{region 'Documentation'}
(*!
<summary>Checks non-overlapping BYTE/WORD array token counts and independent array bounds.</summary>
<description>
Adjacent tokens count separately; overlapping candidates do not share elements.
Word patterns deliberately contain equal low bytes with different high bytes.
Oversized tokens and empty selected ranges are normal parameter errors, not
manufactured empty arrays or invalid references.
Independent scenarios occupy two calls: bound Reset, then evaluation.
ProcessAssertions checks each call before ProcessTests advances. Literal expected
results belong to SelectScenario, not to a copy of the production comparison.
The local capture is cleared before each call and checked in subject-call order.
FirstFailedScenario and FailedDuringEvaluation retain the first mismatch.
Continuation scenarios explicitly retain the prior subject state. The Test Case
owns all input storage; no invalid or dangling references are constructed.
</description>
*)
{endregion}
FUNCTION_BLOCK Test_AssertionArrayTokenCount EXTENDS TestCaseBase
VAR
    FEqual : AssertArrayTokenCntEqual_Byte;
    FEqualExpectedResult : E_Result;
    FWideEqual : AssertArrayTokenCntEqual_Word;
    FWideEqualExpectedResult : E_Result;
    FNone : AssertNoArrayToken_Byte;
    FNoneExpectedResult : E_Result;
    FWideRange : AssertArrayTokenCntInRange_Word;
    FWideRangeExpectedResult : E_Result;
    FData : ARRAY[-2..3] OF BYTE;
    FDataBefore : ARRAY[-2..3] OF BYTE;
    FWideData : ARRAY[-2..3] OF WORD;
    FWideDataBefore : ARRAY[-2..3] OF WORD;
    FToken : ARRAY[4..5] OF BYTE;
    FTokenBefore : ARRAY[4..5] OF BYTE;
    FWideToken : ARRAY[-5..-4] OF WORD;
    FWideTokenBefore : ARRAY[-5..-4] OF WORD;
    FStartIndex : DINT;
    FLength : USINT;
    FExpected : UINT;
    FMinimum : UINT;
    FMaximum : UINT;
    FSubjectEnable : BOOL;
    FContinueScenario : BOOL;
    FEqualExpectedFinding : BOOL;
    FEqualExpectedCount : UINT;
    FWideEqualExpectedFinding : BOOL;
    FWideEqualExpectedCount : UINT;
    FNoneExpectedFinding : BOOL;
    FNoneExpectedCount : UINT;
    FWideRangeExpectedFinding : BOOL;
    FWideRangeExpectedCount : UINT;
    FCapture : EventBuffer;
    FEvents : ARRAY[1..CaptureLength] OF ST_Event;
    FCaptureFifo : ST_FifoStatus;
    FCaptureStatus : ST_EventBufferStatus;
    FSetupValid : BOOL;
    FScenario : UINT;
    FChecked : BOOL;
    FEvaluateSubjects : BOOL;
    FObservationReady : BOOL;
    FFirstFailedScenario : UINT;
    FFailedDuringEvaluation : BOOL;
    FResultsMatch : BOOL;
    FResults : AssertTrue;
    FActivityMatch : BOOL;
    FActivity : AssertTrue;
    FInputsMatch : BOOL;
    FInputs : AssertTrue;
    FFindingsMatch : BOOL;
    FFindings : AssertTrue;
END_VAR
VAR CONSTANT
    CaptureLength : UINT := 8;
    ScenarioAdjacentTokens : UINT := 1;
    ScenarioNonOverlapping : UINT := 2;
    ScenarioTrailingPartial : UINT := 3;
    ScenarioLastCandidate : UINT := 4;
    ScenarioAbsent : UINT := 5;
    ScenarioCountMismatch : UINT := 6;
    ScenarioTokenTooLong : UINT := 7;
    ScenarioEmptyRange : UINT := 8;
    ScenarioRangePastEnd : UINT := 9;
    LastScenario : UINT := ScenarioRangePastEnd;
END_VAR

SUPER^();

{region 'Documentation'}
(*!
<summary>Aggregates only outer checks, not intentionally failing subjects.</summary>
*)
{endregion}
METHOD PROTECTED AggregateResults
VAR_INPUT
    Aggregator : I_ResultAggregator; //! Borrowed result sink owned by the outer Test Case; add this test's checking Assertions without resetting or retaining the sink.
END_VAR
Aggregator.AddProvider(Provider := FResults);
Aggregator.AddProvider(Provider := FActivity);
Aggregator.AddProvider(Provider := FInputs);
Aggregator.AddProvider(Provider := FFindings);
END_METHOD

{region 'Documentation'}
(*!
<summary>Calls each inherited production subject once with caller-owned input storage.</summary>
*)
{endregion}
METHOD PRIVATE CallSubjects
FEqual(Enable := FSubjectEnable,
    State := E_State.Running,
    StartIndex := FStartIndex,
    Length := FLength,
    Expected := FExpected,
    IN := FData,
    Token := FToken);
FWideEqual(Enable := FSubjectEnable,
    State := E_State.Running,
    StartIndex := FStartIndex,
    Length := FLength,
    Expected := FExpected,
    IN := FWideData,
    Token := FWideToken);
FNone(Enable := FSubjectEnable,
    State := E_State.Running,
    StartIndex := FStartIndex,
    Length := FLength,
    IN := FData,
    Token := FToken);
FWideRange(Enable := FSubjectEnable,
    State := E_State.Running,
    StartIndex := FStartIndex,
    Length := FLength,
    Minimum := FMinimum,
    Maximum := FMaximum,
    IN := FWideData,
    Token := FWideToken);
END_METHOD

{region 'Documentation'}
(*!
<summary>Checks one subject finding in call order; expected outcomes come from the scenario.</summary>
*)
{endregion}
METHOD PRIVATE CheckFinding : BOOL //! TRUE when the required finding checks pass; calls requiring no finding also succeed.
VAR_INPUT
    Subject : I_Assertion; //! Assertion interface supplying the expected finding identity.
    ExpectedResult : E_Result; //! Independently authored result expected in the captured finding.
    ExpectedFinding : BOOL; //! TRUE when this scenario requires a finding during active evaluation.
END_VAR
VAR_IN_OUT
    Index : UINT; //! One-based next finding index; advanced when this call checks a required finding.
END_VAR
CheckFinding := TRUE;
IF FEvaluateSubjects AND ExpectedFinding THEN
    CheckFinding := (FEvents[Index].SequenceId = UINT_TO_UDINT(Index))
        AND (FEvents[Index].Name = Subject.Name)
        AND (FEvents[Index].OwnerScope = E_OwnerScope.Assertion)
        AND (FEvents[Index].EventType = E_EventType.Result)
        AND (FEvents[Index].State = E_State.Running)
        AND (FEvents[Index].Result = ExpectedResult)
        AND (FEvents[Index].Message <> '');
    Index := Index + 1;
END_IF;
END_METHOD

{region 'Documentation'}
(*!
<summary>Checks exact finding count and identities; at most one finding per subject.</summary>
*)
{endregion}
METHOD PRIVATE CheckFindings
VAR
    Index : UINT;
    Matches : BOOL;
END_VAR
Index := 1;
FFindingsMatch := TRUE;
Matches := CheckFinding(Subject := FEqual,
    ExpectedResult := FEqualExpectedResult,
    ExpectedFinding := FEqualExpectedFinding,
    Index := Index);
FFindingsMatch := FFindingsMatch AND Matches;
Matches := CheckFinding(Subject := FWideEqual,
    ExpectedResult := FWideEqualExpectedResult,
    ExpectedFinding := FWideEqualExpectedFinding,
    Index := Index);
FFindingsMatch := FFindingsMatch AND Matches;
Matches := CheckFinding(Subject := FNone,
    ExpectedResult := FNoneExpectedResult,
    ExpectedFinding := FNoneExpectedFinding,
    Index := Index);
FFindingsMatch := FFindingsMatch AND Matches;
Matches := CheckFinding(Subject := FWideRange,
    ExpectedResult := FWideRangeExpectedResult,
    ExpectedFinding := FWideRangeExpectedFinding,
    Index := Index);
FFindingsMatch := FFindingsMatch AND Matches;
FFindingsMatch := FFindingsMatch
    AND (FCaptureStatus.SequenceId = UINT_TO_UDINT(Index - 1))
    AND (FCaptureStatus.LostEventCount = 0);
IF FEvaluateSubjects AND (FScenario = ScenarioCountMismatch) THEN
    // SA0175: Fixed byte-substring checks of bounded diagnostic messages; no character offsets.
    {analysis -175}
    FFindingsMatch := FFindingsMatch
        AND (FIND(FEvents[1].Message, 'Actual = 2') > 0)
        AND (FIND(FEvents[4].Message, 'Actual = 2') > 0);
    {analysis +175}
END_IF;
END_METHOD

{region 'Documentation'}
(*!
<summary>Rejects incomplete subject, capture or outer Assertion setup.</summary>
*)
{endregion}
METHOD PROTECTED CheckInitialization : BOOL //! TRUE when the inherited initialization check and this concrete fixture check both accept the setup.
CheckInitialization := SUPER^.CheckInitialization();
IF NOT CheckInitialization THEN
    RETURN;
END_IF;

CheckInitialization := FSetupValid
    AND FResults.IsInitialized
    AND FActivity.IsInitialized
    AND FInputs.IsInitialized
    AND FFindings.IsInitialized;
IF NOT CheckInitialization THEN
    EventPublisher.PublishEvent(Event := CreateFrameworkEvent(Name := Name,
        ResourceName := '',
        State := State,
        Severity := E_EventSeverity.Error,
        Message := 'Text selftest setup failed.'));
END_IF;
END_METHOD

{region 'Documentation'}
(*!
<summary>Checks literal evaluation results, or NotEvaluated on the reset call.</summary>
*)
{endregion}
METHOD PRIVATE CheckResults
IF FEvaluateSubjects THEN
    FResultsMatch := (FEqual.Result = FEqualExpectedResult)
        AND (FWideEqual.Result = FWideEqualExpectedResult)
        AND (FNone.Result = FNoneExpectedResult)
        AND (FWideRange.Result = FWideRangeExpectedResult);
ELSE
    FResultsMatch := (FEqual.Result = E_Result.NotEvaluated)
        AND (FWideEqual.Result = E_Result.NotEvaluated)
        AND (FNone.Result = E_Result.NotEvaluated)
        AND (FWideRange.Result = E_Result.NotEvaluated);
END_IF;
FActivityMatch := (FEqual.Enabled = FSubjectEnable)
    AND (FEqual.ObservationActive = (FEvaluateSubjects AND FSubjectEnable))
    AND (FEqual.EvaluationActive = (FEvaluateSubjects AND FSubjectEnable))
    AND (FWideEqual.Enabled = FSubjectEnable)
    AND (FWideEqual.ObservationActive = (FEvaluateSubjects AND FSubjectEnable))
    AND (FWideEqual.EvaluationActive = (FEvaluateSubjects AND FSubjectEnable))
    AND (FNone.Enabled = FSubjectEnable)
    AND (FNone.ObservationActive = (FEvaluateSubjects AND FSubjectEnable))
    AND (FNone.EvaluationActive = (FEvaluateSubjects AND FSubjectEnable))
    AND (FWideRange.Enabled = FSubjectEnable)
    AND (FWideRange.ObservationActive = (FEvaluateSubjects AND FSubjectEnable))
    AND (FWideRange.EvaluationActive = (FEvaluateSubjects AND FSubjectEnable));
IF FEvaluateSubjects THEN
    FResultsMatch := FResultsMatch
        AND (FEqual.TokenCount = FEqualExpectedCount)
        AND (FWideEqual.TokenCount = FWideEqualExpectedCount)
        AND (FNone.TokenCount = FNoneExpectedCount)
        AND (FWideRange.TokenCount = FWideRangeExpectedCount);
ELSE
    FResultsMatch := FResultsMatch
        AND (FEqual.TokenCount = 0)
        AND (FWideEqual.TokenCount = 0)
        AND (FNone.TokenCount = 0)
        AND (FWideRange.TokenCount = 0);
END_IF;
END_METHOD

{region 'Documentation'}
(*!
<summary>Initializes outer checks and isolates intentional subject findings.</summary>
*)
{endregion}
METHOD PROTECTED Configure
VAR
    Initialized : BOOL;
END_VAR
FPreparationStateCount := 0;
FTestStateCount := 1;
FResults.Initialize(Parent := THIS^,
    AssertionName := 'Results');
FActivity.Initialize(Parent := THIS^,
    AssertionName := 'Activity');
FInputs.Initialize(Parent := THIS^,
    AssertionName := 'Inputs');
FFindings.Initialize(Parent := THIS^,
    AssertionName := 'Findings');
FSetupValid := FCapture.Initialize(Buffer := FEvents,
    FifoControl := FCaptureFifo,
    Status := FCaptureStatus);
FEqual.BindPublisher(Publisher := FCapture);
Initialized := FEqual.Initialize(Parent := THIS^,
    AssertionName := 'Equal');
FSetupValid := FSetupValid AND Initialized;
FWideEqual.BindPublisher(Publisher := FCapture);
Initialized := FWideEqual.Initialize(Parent := THIS^,
    AssertionName := 'WideEqual');
FSetupValid := FSetupValid AND Initialized;
FNone.BindPublisher(Publisher := FCapture);
Initialized := FNone.Initialize(Parent := THIS^,
    AssertionName := 'None');
FSetupValid := FSetupValid AND Initialized;
FWideRange.BindPublisher(Publisher := FCapture);
Initialized := FWideRange.Initialize(Parent := THIS^,
    AssertionName := 'WideRange');
FSetupValid := FSetupValid AND Initialized;
END_METHOD

{region 'Documentation'}
(*!
<summary>Completes abort; no asynchronous resource is owned.</summary>
*)
{endregion}
METHOD PROTECTED ProcessAbort
VAR_INPUT
    Enable : BOOL; //! Phase permission supplied by the owning Test Case; FALSE does not authorize progression, while observation may continue.
END_VAR
IF Enable THEN
    CompleteAbort();
END_IF;
END_METHOD

{region 'Documentation'}
(*!
<summary>Latches this call's checks before progression is permitted.</summary>
*)
{endregion}
METHOD PROTECTED ProcessAssertions
VAR_INPUT
    Enable : BOOL; //! Phase permission supplied by the owning Test Case; FALSE does not authorize progression, while observation may continue.
END_VAR
VAR
    Check : BOOL;
END_VAR
Check := Enable AND FObservationReady;
FResults(Enable := Check,
    State := State,
    IN := FResultsMatch);
FActivity(Enable := Check,
    State := State,
    IN := FActivityMatch);
FInputs(Enable := Check,
    State := State,
    IN := FInputsMatch);
FFindings(Enable := Check,
    State := State,
    IN := FFindingsMatch);
IF Check THEN
    FChecked := TRUE;
END_IF;
END_METHOD

{region 'Documentation'}
(*!
<summary>No Preparation phase is needed.</summary>
*)
{endregion}
METHOD PROTECTED ProcessPreparations
VAR_INPUT
    // SA0033: Required hook; this test has no Preparation phase.
    {attribute 'analysis' := '-33'}
    Enable : BOOL; //! Phase permission supplied by the owning Test Case; FALSE does not authorize progression, while observation may continue.
END_VAR
END_METHOD

{region 'Documentation'}
(*!
<summary>Restarts the scenario sequence and outer checks.</summary>
*)
{endregion}
METHOD PROTECTED ProcessReset
FScenario := ScenarioAdjacentTokens;
FChecked := FALSE;
FSubjectEnable := FALSE;
FContinueScenario := FALSE;
FEvaluateSubjects := FALSE;
FObservationReady := FALSE;
FFirstFailedScenario := 0;
FFailedDuringEvaluation := FALSE;
FCapture.Reset();
ResetSubjects();
FResults.Reset();
FActivity.Reset();
FInputs.Reset();
FFindings.Reset();
CompleteReset();
END_METHOD

{region 'Documentation'}
(*!
<summary>Consumes reset before each independent scenario; continuation retains subject state.</summary>
*)
{endregion}
METHOD PROTECTED ProcessTests
VAR_INPUT
    Enable : BOOL; //! Phase permission supplied by the owning Test Case; FALSE does not authorize progression, while observation may continue.
END_VAR
IF NOT Enable THEN
    RETURN;
END_IF;

IF FChecked THEN
    FChecked := FALSE;
    FObservationReady := FALSE;
    IF FEvaluateSubjects THEN
        IF FScenario = LastScenario THEN
            CompleteTests();
            RETURN;
        END_IF;
        FScenario := FScenario + 1;
    END_IF;
    FEvaluateSubjects := NOT FEvaluateSubjects;
END_IF;

IF NOT SelectScenario() THEN
    RETURN;
END_IF;
IF FContinueScenario THEN
    FEvaluateSubjects := TRUE;
END_IF;
FCapture.Reset();
IF NOT FEvaluateSubjects THEN
    ResetSubjects();
END_IF;
FDataBefore := FData;
FWideDataBefore := FWideData;
FTokenBefore := FToken;
FWideTokenBefore := FWideToken;
CallSubjects();
CheckResults();
FInputsMatch := (FData[-2] = FDataBefore[-2])
    AND (FData[-1] = FDataBefore[-1])
    AND (FData[0] = FDataBefore[0])
    AND (FData[1] = FDataBefore[1])
    AND (FData[2] = FDataBefore[2])
    AND (FData[3] = FDataBefore[3])
    AND (FWideData[-2] = FWideDataBefore[-2])
    AND (FWideData[-1] = FWideDataBefore[-1])
    AND (FWideData[0] = FWideDataBefore[0])
    AND (FWideData[1] = FWideDataBefore[1])
    AND (FWideData[2] = FWideDataBefore[2])
    AND (FWideData[3] = FWideDataBefore[3])
    AND (FToken[4] = FTokenBefore[4])
    AND (FToken[5] = FTokenBefore[5])
    AND (FWideToken[-5] = FWideTokenBefore[-5])
    AND (FWideToken[-4] = FWideTokenBefore[-4]);
CheckFindings();
IF (FFirstFailedScenario = 0)
    AND NOT (FResultsMatch AND FActivityMatch AND FInputsMatch AND FFindingsMatch) THEN
    FFirstFailedScenario := FScenario;
    FFailedDuringEvaluation := FEvaluateSubjects;
END_IF;
FObservationReady := TRUE;
END_METHOD

{region 'Documentation'}
(*!
<summary>Queues reset; the next bound FB call consumes it without evaluating.</summary>
*)
{endregion}
METHOD PRIVATE ResetSubjects
FEqual.Reset();
FWideEqual.Reset();
FNone.Reset();
FWideRange.Reset();
END_METHOD

{region 'Documentation'}
(*!
<summary>Selects explicit stimuli and expected results for one scenario.</summary>
*)
{endregion}
METHOD PRIVATE SelectScenario : BOOL //! TRUE after selecting a supported scenario and its literal expectations; FALSE reports an unknown scenario.
SelectScenario := FALSE;
FSubjectEnable := TRUE;
FContinueScenario := FALSE;
FData[-2] := 1;
FData[-1] := 2;
FData[0] := 1;
FData[1] := 2;
FData[2] := 9;
FData[3] := 9;
FWideData[-2] := WORD#16#0101;
FWideData[-1] := WORD#16#0202;
FWideData[0] := WORD#16#0101;
FWideData[1] := WORD#16#0202;
FWideData[2] := 1;
FWideData[3] := 2;
FToken[4] := 1;
FToken[5] := 2;
FWideToken[-5] := WORD#16#0101;
FWideToken[-4] := WORD#16#0202;
FStartIndex := -2;
FLength := 6;
FExpected := 2;
FMinimum := 2;
FMaximum := 2;
CASE FScenario OF
    ScenarioAdjacentTokens:
        FEqualExpectedResult := E_Result.Passed;
        FEqualExpectedFinding := FALSE;
        FEqualExpectedCount := 2;
        FWideEqualExpectedResult := E_Result.Passed;
        FWideEqualExpectedFinding := FALSE;
        FWideEqualExpectedCount := 2;
        FNoneExpectedResult := E_Result.Failed;
        FNoneExpectedFinding := TRUE;
        FNoneExpectedCount := 2;
        FWideRangeExpectedResult := E_Result.Passed;
        FWideRangeExpectedFinding := FALSE;
        FWideRangeExpectedCount := 2;
    ScenarioNonOverlapping:
        FLength := 3;
        FData[-1] := 1;
        FToken[5] := 1;
        FWideData[-1] := WORD#16#0101;
        FWideToken[-4] := WORD#16#0101;
        FExpected := 1;
        FMinimum := 1;
        FMaximum := 1;
        FEqualExpectedResult := E_Result.Passed;
        FEqualExpectedFinding := FALSE;
        FEqualExpectedCount := 1;
        FWideEqualExpectedResult := E_Result.Passed;
        FWideEqualExpectedFinding := FALSE;
        FWideEqualExpectedCount := 1;
        FNoneExpectedResult := E_Result.Failed;
        FNoneExpectedFinding := TRUE;
        FNoneExpectedCount := 1;
        FWideRangeExpectedResult := E_Result.Passed;
        FWideRangeExpectedFinding := FALSE;
        FWideRangeExpectedCount := 1;
    ScenarioTrailingPartial:
        FLength := 3;
        FExpected := 1;
        FMinimum := 1;
        FMaximum := 1;
        FEqualExpectedResult := E_Result.Passed;
        FEqualExpectedFinding := FALSE;
        FEqualExpectedCount := 1;
        FWideEqualExpectedResult := E_Result.Passed;
        FWideEqualExpectedFinding := FALSE;
        FWideEqualExpectedCount := 1;
        FNoneExpectedResult := E_Result.Failed;
        FNoneExpectedFinding := TRUE;
        FNoneExpectedCount := 1;
        FWideRangeExpectedResult := E_Result.Passed;
        FWideRangeExpectedFinding := FALSE;
        FWideRangeExpectedCount := 1;
    ScenarioLastCandidate:
        FStartIndex := -1;
        FLength := 3;
        FExpected := 1;
        FMinimum := 1;
        FMaximum := 1;
        FEqualExpectedResult := E_Result.Passed;
        FEqualExpectedFinding := FALSE;
        FEqualExpectedCount := 1;
        FWideEqualExpectedResult := E_Result.Passed;
        FWideEqualExpectedFinding := FALSE;
        FWideEqualExpectedCount := 1;
        FNoneExpectedResult := E_Result.Failed;
        FNoneExpectedFinding := TRUE;
        FNoneExpectedCount := 1;
        FWideRangeExpectedResult := E_Result.Passed;
        FWideRangeExpectedFinding := FALSE;
        FWideRangeExpectedCount := 1;
    ScenarioAbsent:
        FToken[4] := 7;
        FWideToken[-5] := 7;
        FExpected := 0;
        FMinimum := 0;
        FMaximum := 0;
        FEqualExpectedResult := E_Result.Passed;
        FEqualExpectedFinding := FALSE;
        FEqualExpectedCount := 0;
        FWideEqualExpectedResult := E_Result.Passed;
        FWideEqualExpectedFinding := FALSE;
        FWideEqualExpectedCount := 0;
        FNoneExpectedResult := E_Result.Passed;
        FNoneExpectedFinding := FALSE;
        FNoneExpectedCount := 0;
        FWideRangeExpectedResult := E_Result.Passed;
        FWideRangeExpectedFinding := FALSE;
        FWideRangeExpectedCount := 0;
    ScenarioCountMismatch:
        FExpected := 1;
        FMinimum := 3;
        FMaximum := 4;
        FEqualExpectedResult := E_Result.Failed;
        FEqualExpectedFinding := TRUE;
        FEqualExpectedCount := 2;
        FWideEqualExpectedResult := E_Result.Failed;
        FWideEqualExpectedFinding := TRUE;
        FWideEqualExpectedCount := 2;
        FNoneExpectedResult := E_Result.Failed;
        FNoneExpectedFinding := TRUE;
        FNoneExpectedCount := 2;
        FWideRangeExpectedResult := E_Result.Failed;
        FWideRangeExpectedFinding := TRUE;
        FWideRangeExpectedCount := 2;
    ScenarioTokenTooLong:
        FLength := 1;
        FEqualExpectedResult := E_Result.Error;
        FEqualExpectedFinding := TRUE;
        FEqualExpectedCount := 0;
        FWideEqualExpectedResult := E_Result.Error;
        FWideEqualExpectedFinding := TRUE;
        FWideEqualExpectedCount := 0;
        FNoneExpectedResult := E_Result.Error;
        FNoneExpectedFinding := TRUE;
        FNoneExpectedCount := 0;
        FWideRangeExpectedResult := E_Result.Error;
        FWideRangeExpectedFinding := TRUE;
        FWideRangeExpectedCount := 0;
    ScenarioEmptyRange:
        FLength := 0;
        FEqualExpectedResult := E_Result.Error;
        FEqualExpectedFinding := TRUE;
        FEqualExpectedCount := 0;
        FWideEqualExpectedResult := E_Result.Error;
        FWideEqualExpectedFinding := TRUE;
        FWideEqualExpectedCount := 0;
        FNoneExpectedResult := E_Result.Error;
        FNoneExpectedFinding := TRUE;
        FNoneExpectedCount := 0;
        FWideRangeExpectedResult := E_Result.Error;
        FWideRangeExpectedFinding := TRUE;
        FWideRangeExpectedCount := 0;
    ScenarioRangePastEnd:
        FStartIndex := 3;
        FLength := 2;
        FEqualExpectedResult := E_Result.Error;
        FEqualExpectedFinding := TRUE;
        FEqualExpectedCount := 0;
        FWideEqualExpectedResult := E_Result.Error;
        FWideEqualExpectedFinding := TRUE;
        FWideEqualExpectedCount := 0;
        FNoneExpectedResult := E_Result.Error;
        FNoneExpectedFinding := TRUE;
        FNoneExpectedCount := 0;
        FWideRangeExpectedResult := E_Result.Error;
        FWideRangeExpectedFinding := TRUE;
        FWideRangeExpectedCount := 0;
ELSE
    Error(Message := 'Unknown Assertion scenario.');
    RETURN;
END_CASE;
SelectScenario := TRUE;
END_METHOD

END_FUNCTION_BLOCK

(* stored: Version 1.1.0.1
   POU Test_AssertionArrayTokenCount: Id {a869522e-5487-4e1a-921d-4fd4cab0694f}, SpecialFunc None
   Folder Internal: Id {3642be2a-c7c5-4817-a3d0-515a984b274a}
   Method AggregateResults: Id {3ccffe37-f0c7-4a2e-86ea-2892f2032958}
   Method CallSubjects: Id {349bf756-2bf6-4b57-a665-f977aacbf492}
   Method CheckFinding: Id {278c8903-5a40-4983-9d44-a41f820fda91}
   Method CheckFindings: Id {2f80efa3-daca-481d-9fe6-441653bd06b8}
   Method CheckInitialization: Id {020c46ec-0638-4d9b-85fc-4bd233aefc44}
   Method CheckResults: Id {af25168c-4b1c-4c30-9712-b55e66b125d8}
   Method Configure: Id {f9fcc5fa-61c5-45cf-b012-e00baf48d255}
   Method ProcessAbort: Id {874f4ea2-8126-4c39-8c16-1b2cc5b219c1}
   Method ProcessAssertions: Id {163713b6-19ea-4d05-b995-589f30aa7346}
   Method ProcessPreparations: Id {1c17ad36-bb5d-4c5f-8468-d3bec19da919}
   Method ProcessReset: Id {d166470d-1fdc-42c4-9dc5-82037a5e8c12}
   Method ProcessTests: Id {b0de9e74-163e-4071-943d-a01d7d604252}
   Method ResetSubjects: Id {221f7488-f606-41ab-8d15-86755a9cfb33}
   Method SelectScenario: Id {1158dc19-5014-4ffb-add1-c485135f94dd} *)
